Fanuc KAREL source: kt00859.KL

-- PROVISIONAL review KL for V940-1; original PC SHA256 4aa34fe178cab1bc00ac9dc3057f31129e1a6864e89b89c49238311f223f0da2
-- Incomplete behavior may be omitted. Consult companion uncertainty JSON. Do not deploy.
PROGRAM KT00859
%NOLOCKGROUP
VAR
  R1 : REAL
  R2 : REAL
  OUT : REAL
BEGIN
  -- V9_ZERO_TABLE_METADATA_HINT layout=0001; no indexed target words; source/name/runtime held
  -- UNRESOLVED_PC offsets 5-16; opcodes 2E,23
  -- UNRESOLVED_PC offsets 21-32; opcodes 2E,23
  -- UNRESOLVED_PC offsets 37-48; opcodes 2E,23
  -- UNRESOLVED_PC offsets 53-64; opcodes 2E,23
  -- UNRESOLVED_PC offsets 69-85; opcodes 27,22,76,64,23
  -- UNRESOLVED_PC offsets 90-94; opcodes 7F
END KT00859
